Staubli VAL3: simulateTRAJ.pgx

public program simulateTRAJ(string x_sKey)
  local bool l_bResult
begin
  if !rs:bIsCycle and workingMode()==1
    l_bResult=userPageConfirm("是否模拟TRAJ："+x_sKey+"？")
    if l_bResult
      resetMotion()
      rs:bSimulate=true
      rs:bGOTO=false
      //添加traj任务‘
      taskCreate "simulate",100,trajectory:makeTraj(x_sKey)
      //
      sMsg="模拟TRAJ过程。。。"
      sMsg=rs:sTrajStatus
      call simulate_UI()
    endIf
  else
    userPageAlert("条件不满足：不再生产周期&切换到手动模式")
  endIf
end
